(* IEC 61131-3 sources: PLC-Static-Analysis/modules/plc-rules/src/test/resources/PLCA-L017, 2 files *)

(* ---- compliant.st ---- *)
PROGRAM P_L017ok
VAR
    n : INT;
    m : INT;
    r : REAL;
    b : BOOL;
    c : BOOL;
    q : BOOL;
END_VAR
IF b THEN
    RETURN;
END_IF
q := TRUE;
IF b THEN
    q := FALSE;
ELSIF c THEN
    RETURN;
ELSE
    m := 1;
END_IF
END_PROGRAM

(* ---- noncompliant.st ---- *)
PROGRAM P_L017
VAR
    n : INT;
    m : INT;
    r : REAL;
    b : BOOL;
    c : BOOL;
    q : BOOL;
END_VAR
IF b THEN
    RETURN;
ELSE // PLCA-L017
    q := TRUE;
END_IF
FOR n := 1 TO 10 DO
    IF b THEN
        q := TRUE;
        CONTINUE;
    ELSIF c THEN
        EXIT;
    ELSE // PLCA-L017
        m := n;
    END_IF
END_FOR
END_PROGRAM
